Fanuc KAREL source: KT00218.KL

PROGRAM KT00218
%NOLOCKGROUP
VAR
  H1: ARRAY[2] OF SHORT
  B2: BOOLEAN
  OUT: INTEGER
BEGIN
  H1[1] = 2
    B2 = FALSE
  OUT = H1[1] AND B2
END KT00218
